// TIA Portal V20 export
Screen "Call_ServiceButtons"  1276x673
  ScreenItem "Title_OPMode1_ScreenOverview_X390_Y2" at 5,7 size 1262x30  Type=HmiTextBox
  ScreenItem "Faceplate container_5" at 0,33 size 622x206  Type=HmiFaceplateContainer
  ScreenItem "Text box_5" at 0,0 size 622x30  Type=HmiTextBox
  ScreenItem "Faceplate container_7" at 0,33 size 622x206  Type=HmiFaceplateContainer
  ScreenItem "Text box_7" at 0,0 size 622x30  Type=HmiTextBox
  ScreenItem "Faceplate container_8" at 0,33 size 622x206  Type=HmiFaceplateContainer
  ScreenItem "Text box_8" at 0,0 size 622x30  Type=HmiTextBox
  ScreenItem "Faceplate container_1" at 5,73 size 619x179  Type=HmiFaceplateContainer
  ScreenItem "Text box_1" at 5,40 size 622x30  Type=HmiTextBox
  ScreenItem "Faceplate container_2" at 645,73 size 619x179  Type=HmiFaceplateContainer
  ScreenItem "Text box_2" at 645,40 size 622x30  Type=HmiTextBox
  ScreenItem "Faceplate container_3" at 5,285 size 619x179  Type=HmiFaceplateContainer
  ScreenItem "Text box_3" at 5,252 size 622x30  Type=HmiTextBox
  ScreenItem "Faceplate container_4" at 645,285 size 619x179  Type=HmiFaceplateContainer
  ScreenItem "Text box_4" at 645,252 size 622x30  Type=HmiTextBox
  ScreenItem "Button_15" at 1170,8 size 98x31  Type=HmiButton
  ScreenItem "Faceplate container_6" at 5,496 size 619x179  Type=HmiFaceplateContainer
  ScreenItem "Text box_6" at 5,463 size 622x30  Type=HmiTextBox
  ScreenItem "Faceplate container_9" at 645,496 size 619x179  Type=HmiFaceplateContainer
  ScreenItem "Text box_9" at 645,463 size 622x30  Type=HmiTextBox
